TYPE "ST_AirPressureDevice"
VERSION : 0.1
   STRUCT
      Conflicting : Bool;
      Contradictory : Bool;
      ConflictSinceMs : UDInt;
   END_STRUCT;

END_TYPE

